Staubli VAL3: onStart.pgx

program onStart()
  local num l_i
  local num l_nResult
begin
  call saveData:setBaseJOG(saveData:nJogTool)
  sToolIndex=toString("",saveData:nJogTool)
  sSelZone=""
  sLastZone=""
  resize(sList,1,size(safeTemp:zZoneItem))

  for l_i = 0 to size(sList)-1
    sList[l_i]=toString("",l_i)+","+safeTemp:zZoneItem[l_i].sID
  endFor
  bActive=false
  for l_i = 0 to 5
    nFrame[l_i]=0
    nTRSF1[l_i]=0
    nTRSF2[l_i]=0
  endFor
end
